(* IEC 61131-3 sources: Caravan/Archiv/12-04-19/Stations/MachineControl/MachineControl/Network/HW_Network, 1 file *)

(* ---- ONE_HW_Network_Table.st ---- *)
#define OBJECTS_CONFIG

//Define part of class SdiasBase
//Address to access the Dataobject list via SPI SDO Read
#define SDIAS_SPI_DATA_OBJECT_LIST_PAGE_ADDRESS 16#FFFF
#define SDIAS_SPI_DATA_OBJECT_LIST_PAGE_OFFSET 16#00
#define SDIAS_SPI_DATA_OBJECT_LIST_IDENTIFIER 16#12345678

//Defines the number of optional list elements in the SPI List

#define SDIAS_SPI_NUMBER_OF_OPTIONAL_ELEMENTS 7

//#pragma message("EisMic 27.06.2014 14:44 \ Noch schauen ob ichs besser machen kann")
#define SDIAS_SPI_HEADER_BEFORE_OPTIONAL_ELEMENTS 16#18
#define SDIAS_SPI_HARDWARE_VERSION_OFFSET 16#C
#define SDIAS_SPI_VENDOR_ID_OFFSET 16#0

//SPI List IDs
#define SDIAS_SPI_IDENTIFICATION_LIST_ID 1
#define SDIAS_SPI_FLASH_CONFIGURATION_ID 2
#define SDIAS_SPI_VENDOR_NAME_ID 3
#define SDIAS_SPI_DEVICE_NAME_ID 4
#define SDIAS_SPI_SERIAL_NUMBER_ID 5
#define SDIAS_SPI_ORDERING_NUMBER_ID 6
#define SDIAS_SPI_DOCUMENTATION_PDF_ID 7
#define SDIAS_SPI_CALIB_DATA_ID 10
#define SDIAS_SPI_PDO_INFORMATION_ID 128
#include "..\..\Class\SdiasManager\SdiasManager.h"
#include "..\..\Class\SdiasBase\SdiasBase.h"
#include "..\..\Class\HwControl\HwControl.h"
#include "..\..\Source\interfaces\lsl_st_hardwaretree.h"
#include "..\..\Source\interfaces\lsl_st_mt.h"
//Define part of class AI075
#define DEVICE_ID_AI075 1007

#define AI075_ADDR_CYC_WRITE        16#000
#define AI075_ADDR_CYC_READ         16#080
#define AI075_ADDR_CFG_FIRMWARE     16#100
#define AI075_ADDR_STATE_FIRMWARE   16#180

#define AI075_SDO_RESPONSE_TIMEOUT  SDIAS_SDO_TIMEOUT * 2

#define AI075_LENGTH_STATE_FIRMWARE 2
#define AI075_NUMBER_OF_ANALOG_IN   6
#define AI075_NUMBER_OF_TMP_IN      1
#define AI075_INVALID_VALUE         16#80000010$DINT
#define AI075_CABLE_BREAK_MASK      16#7F  //7 BITS
#define AI075_SHORT_CIRCUIT_MASK    16#03  //2 BITS
#define AI075_SAMPLE_POINT_MASK     16#0F  //4 BITS
#define AI075_OFFSET_SAMPLE_POINT_BITS 11

#define AI075_FIRMWARE_MIN          -10000
#define AI075_FIRMWARE_MAX          10000

//Sample Point Defines
//**************************************************************
#define AI075_FIRMWARE_VERSION_SAMPLE_POINTS_AVAILABLE  16#200
#define AI075_SAMPLE_POINTS_OFFSET_AFTER_SYNC   15    //Minimal offset that a sample point can be set after sync
#define AI075_SAMPLE_POINTS_OFFSET_BEFORE_SYNC  162   //Maximal offset that a sample point can be before next sync
//Define part of class AI088
#define DEVICE_ID_AI088 1009

#define AI088_ADDR_CYC_WRITE        16#000
#define AI088_ADDR_CYC_READ         16#080
#define AI088_ADDR_CFG_FIRMWARE     16#100
#define AI088_ADDR_STATE_FIRMWARE   16#180

#define AI088_SDO_RESPONSE_TIMEOUT  SDIAS_SDO_TIMEOUT * 2

#define AI088_LENGTH_STATE_FIRMWARE 2
#define AI088_NUMBER_OF_TMP_INPUT   10
#define AI088_CABLE_BREAK_MASK      16#3FF  //10 BITS
#define AI088_SHORT_CIRCUIT_MASK    16#3    //2 BITS
#define AI088_INVALID_VALUE         16#80000010$DINT

#define AI088_FIRMWARE_VERSION_INT_TEMP_REF 16#200  //Firmware version since when internal temperature reference and message counter are supported
#define AI088_HARDWARE_VERSION_INT_TEMP_REF 16#300  //Hardware version since when internal temperature reference are supported
// for TMP_XSelect = 10: data coming from FW may be originally negative but are
// sent as UINT type - so negativ values are sent as very big UINT values
// values greater than AI088_THRESHOLD_NEG_VALS are interpreted as neative ones
#define AI088_THRESHOLD_NEG_VALS  59000
#define AI088_SUBTRACT_FOR_INT    16#10000
//Define part of class BusInterfaceSDIASInternal
#define BUSIF_INTERNAL_MAX_NR_DO 100

// Defines for Mutex Generation
#define INTERNAL_STR_MUTEX_NAME_SEPERATOR ".."
#define INTERNAL_MUTEX_NAME_END_LENGTH 5
#define INTERNAL_MUTEX_NAME_MAX_LENGTH 32
#include "..\..\Source\BusInterface.h"
//Define part of class DI203
#define DEVICE_ID_DI203 1018
#include "..\..\Class\HwControl\watchdog.h"
#include "..\..\Source\interfaces\lsl_st_sysinfo.h"
#include "..\..\Source\interfaces\lsl_st_systrace.h"
#include <.\lsl_st_mt.h>
//Define part of class SafetyUDP
#define SAFETY_UDP_MAX_SOCKETS                6     // Max number of socket

#define SAFETY_UDP_CLT_SEND_OK                0    // Send ok
#define SAFETY_UDP_CLT_INVALID_HANDLE        -1    // Invalid handle
#define SAFETY_UDP_CLT_NOT_OPEN              -2    // Socket is not open
#define SAFETY_UDP_CLT_SEND_FAILED           -3    // Send failed
#define SAFETY_UDP_CLT_SEND_BUFFER_FULL      -4    // Send buffer is full
#define SAFETY_UDP_CLT_DATA_TO_BIG           -5    // Data to big

#define SAFETY_UDP_MAXIMUM_SEGMENT_SIZE    1452    // Maximum of user data

#define SAFETY_UDP_TIMEOUT_OPENSOCKET    (1000)    //timeout for opening socket

#define SAFETY_UDP_RECEIVE_TIMEOUT          800

#define SAFETY_UDP_TX_BUFFER_SIZE          1024
//Define part of class SafetyManager
#define LogBufferSize 1000
#include "..\..\Class\SafetyManager\SafetyManager.h"
#include "..\..\Source\interfaces\lsl_st_safetydll.h"
//Define part of class SdiasManager
#define SDIAS_SDO_MAX_LENGTH              128
#define SDIAS_SDO_RINGBUFFER_NO            64
#define SDIAS_SDO_CHANNEL_NO                3   // fixed in the VI hardware to be 3

// watchdog trigger interval (after 130ms of no trigger the SDIAS HW goes into reset again and takes at least another 10ms to be ready again)
#define SDIAS_WATCHDOG_TRIGGER_TIME        40

// time needed by sdias modules to start up after the watchdog is triggered the first time in ms
#define SDIAS_HARDWARE_STARTUP_TIME        15

// sdias manager needs 2 ticks to handle event for read task (measure sync time)
#define SDIAS_SYNC_MEASURE_TICKS            2

// after activating the PLL SyncOut it takes 3 cycles until the SDIAS sync can be injected
#define SDIAS_CYCLES_WAIT_AFTER_SYNC_ENABLE 3

// wait 1 bus cycle at start to get valid numbers in the task info
#define SDIAS_TASKINFO_READY_TICKS          1

// time to wait (in ms) until other tasks in the same or lower priority than post init have done their stuff
#define SDIAS_WAIT_TIME_IN_POST_INIT        1

#define SIZE_PER_SDIAS_CLIENT               16#0400

// for far memory accesses: 1 module can hold maximum 256 1K blocks (0-255)
#define SDIAS_1K_BLOCK_NO                       256

// far memory accesses maximum length in bytes
#define SDIAS_MAX_SIZE_FAR_MEM_ACCESS           127

#define SDIAS_OFFSET_HW_CONFIG              16#FF00
#define SDIAS_OFFSET_TASK_EVENT_IDS         16#FF10
#define SDIAS_OFFSET_FEATURE_INFO           16#FF18
#define SDIAS_OFFSET_APPLI_LED_STATES       16#FF20
#define SDIAS_OFFSET_SYNC_INJECTION_CFG     16#FF3D
#define SDIAS_OFFSET_TRIGGER_UNIT_SETUP_0   16#FF41
#define SDIAS_OFFSET_TRIGGER_UNIT_SETUP_1   16#FF45
#define SDIAS_OFFSET_TASK_START_CFG_0       16#FF60
#define SDIAS_OFFSET_TASK_CONFIG_0          16#FF86
#define SDIAS_OFFSET_TASK_CONFIG_1          16#FF96
#define SDIAS_OFFSET_TASK_INFO_1            16#FF94
#define SDIAS_OFFSET_TASK_HANDSHAKE_1       16#FF9B
#define SDIAS_OFFSET_TASK_DURATION_TIME_1   16#FF9C
#define SDIAS_OFFSET_TASK_DURATION_TIME_2   16#FFAC
#define SDIAS_OFFSET_TASK_CONFIG_2          16#FFA6

#define SDIAS_RETRIES_ALLOWED         2

// mask to get global error flag out of message counter byte of SDO responses
#define SDIAS_MASK_GLOBAL_ERROR_FLAG        16#80

// mask to get message counter out of message counter byte of SDO responses
#define SDIAS_MASK_MESSAGE_COUNTER          16#3F

#define SDIAS_EVENT_MASK_ID_SYNC_OUT0       16#10
#define SDIAS_EVENT_MASK_ID_SYNC_OUT1       16#11
#define SDIAS_EVENT_MASK_ID_SYNC_OUT2       16#12
#define SDIAS_EVENT_MASK_ID_SYNC_OUT3       16#13

#define SDIAS_MANAGER_SYNC_SYNCOUT_ID       16#85
#define SDIAS_TASK_START_EVENT_SYNCOUT_ID   16#86

#define SDIAS_PLACE_NO_MODULE_ADDED_SO_FAR  16#80000000

#define SDIAS_TRIGGER_UNIT_BYTE_SIZE        2

#define SDIAS_WAIT_TIME_FIRMWARE_HANDSHAKE  5 * 1000

// if the firmware version is below this, there might be problems with SCP111 and other modules => print warning at startup
#define SDIAS_FW_VERSION_SDO_ERROR_FIXED    16#120

// if the protocol version ist below this, Control Read/Broadcast Write Command is not supported by sdiasmanager
#define SDIAS_PROTOCOLVERSION_BROADCAST     16#120

// if the cil version ist below this, Control Read/Broadcast Write Command is not supported by OS for local SDIAS.
#define SDIAS_CILVERSION_BROADCAST         16#5001

// timeout for blocking the init during initialisation (in ms)
#define SDIAS_INIT_BLOCK_TIMEOUT            20 * 1000

#define SDIAS_MUTEX_NAME_END_LENGTH 3
#define SDIAS_MUTEX_NAME_MAX_LENGTH 32
#define SDIAS_MUTEX_STR_SEPERATOR   ".."

//#define SDIAS_RT_TIME_MEASUREMENT
#ifdef SDIAS_RT_TIME_MEASUREMENT
  #pragma message("ATTENTION: SDIAS real time measurement is active and needs additional ressources in the realtime task")
#endif

(* SDIAS data object commands  *)
#define	 SDIAS_CMD_END							  0x00			(* End command										          *)
#define	 SDIAS_CMD_ACC_MEMORY				  0x01			(* Access dpram memory								      *)
#define	 SDIAS_CMD_ACC_CONTROL				0x02			(* Access dpram control memory						  *)
#define	 SDIAS_CMD_GLOBAL						  0x03			(* SDIAS global command								      *)
#define	 SDIAS_CMD_COPY_LOCAL					0x04			(* DPRAM copy command in local dpram				*)
#define	 SDIAS_CMD_JMP_LOCAL					0x05			(* DPRAM jump command in local dpram 				*)
#define  SDIAS_CMD_ACC_MEMORY_FAR     0x07      (* SDIAS Far Memory Access                  *)

(* SDIAS defines for data object handling *)
// Write data oject list
#define	 SDIAS_DOL_WRITE_USAGE_DOL_EMPTY	  0x20			(* Usage of empty write dol list (wachtdog trigger + end command)   *)
#define	 SDIAS_DOL_WRITE_USAGE_DTA_EMPTY	  0x03			(* Usage of empty write dol data (DO ctrl of 2x copy command for task information + DO ctrl of watchdog trigger      *)
#define	 SDIAS_DOL_WRITE_OFFSET_END_CMD			0x10			(* One data object in list - offset = 1 DO size = 0x10						  *)
#define	 SDIAS_DOL_WRITE_OFFSET_FIRST_DTA		0x02			(* Offset of first data byte of second copy command = 2 (DO ctrl)   *)
#define	 SDIAS_DOL_WRITE_OFFSET_LAST_DTA		0x02			(* Offset of last data byte of second copy command = 2 (DO ctrl )   *)

// Read data oject list
#define	 SDIAS_DOL_READ_USAGE_DOL_EMPTY	    0x30			(* Usage of empty read dol list (2x task info copy command + end command)   *)
#define	 SDIAS_DOL_READ_USAGE_DTA_EMPTY	    0x0D			(* Usage of empty write dol data (DO ctrl of 2x copy command for task information + DO ctrl of watchdog trigger      *)
#define	 SDIAS_DOL_READ_OFFSET_END_CMD			0x20			(* One data object in list - offset = 1 DO size = 0x10						          *)
#define	 SDIAS_DOL_READ_OFFSET_FIRST_DTA		0x07			(* Offset of first data byte of second copy command = 7 = DO state          *)
#define	 SDIAS_DOL_READ_OFFSET_LAST_DTA		  0x0C			(* Offset of last data byte of second copy command = 12 (last byte of task information)       *)

//Versionsnumber where SDIAS SPI Read Accesses are available
#define  SDIAS_SDO_SPI_FIRMWARE_VERSION_AVAILABLE 16#0120

//error info mask
#define  SDIAS_ERROR_INFO_MASK    2#1000011000011111

// Broadcast DO Info
#define SDIAS_OFFSET_CLIENT_CTRLTIMESTAMP   16#0190
#define SDIAS_NR_TIMEBROADCAST_DOS 2
#define SDIAS_TIMEBROADCAST_SUBCMD 16#B0
#include "..\..\Source\interfaces\lsl_st_pll.h"
//Define part of class SdiasPLC
#define SDIASM_OBJECT_PATH            16#88000002   // Object Path for VSDIASmanager Length = 2 (First 2byte), Domain = 0 (3rd byte), Escape Sequence SDIAS (4th byte)
//Define part of class SR020
#define DEVICE_ID_SR020             1015        //DeviceID of SR020

#define SR020_ADDR_CYC_WRITE        16#00       //Address for TPDO
#define SR020_ADDR_CYC_READ         16#0A       //Address for RPDO

#define SR020_ADDR_CFG_FIRMWARE     16#200      //Address-Offset to the Configuration of the Firmware
#define SR020_ADDR_STATE_FIRMWARE   16#280      //Address-Offset to the Status of the Firmware
#define SR020_ADDR_I2T_THRESHOLD    16#20       //Address-Offset to Write I²T Threshold
#define SR020_ADDR_LED_MAX          16#18       //Address-Offset to get LED Configuration-Values

//Define for the H-Brdige
//-----------------------------------------------------------
#define SR020_GATE_A_LOW		          2#0100000000000000    //Bit-Configuration for Enable GateA Low-Switch
#define SR020_GATE_A_HIGH		          2#0001000000000000    //Bit-Configuration for Enable GateA High-Switch
#define SR020_GATE_B_LOW		          2#1000000000000000    //Bit-Configuration for Enable GateB Low-Switch
#define SR020_GATE_B_HIGH		          2#0010000000000000    //Bit-Configuration for Enable GateB High-Switch

#define SR020_MASK_CONTROL	          16#0FFF     //Mask for Output Sequence Bits
#define SR020_MASK_TIME		            16#F000     //Mask for TimeValue

#define SR020_T_SWITCH                41      //Delay Time for Switch
#define SR020_DEFAULT_SEQ_INIT        1       //Initilization for Sequencer => After 1 FPGA-Cycle switch to next Sequency

#define SR020_FPGA_FREQ_MHZ           50    //Frequency of FPGA

#define SR020_SDO_RESPONSE_TIMEOUT  SDIAS_SDO_TIMEOUT * 2     //SDO-Response Timeout

//#define SR020_I2T_THRESHOLD          16000000   //Maximal allowed I²T Value in mA²s ==> 16 A²s
//#pragma message ("TarPet: dieser Wert wurde vorest empirisch ermittelt und sollte noch genau bestimmt werden");
#define SR020_I2T_THRESHOLD          78000   //Maximal allowed I²T Value in mA²s ==> 16 A²s

#define SR020_SPEED_SCALING          10000      //Scaling of the Server Speed (0.00% to 100.00%)
#define SR020_MINPULSE_SCALING       1000       //Scaling of the Server MinPulse (0.0% to 100.0%)

#define SR020_STATUS_BITS_LATCHED  2#0001110011110 // no DC OK info, no sequencer info, no Overtemperature and no I2C error
#define SR020_STATUS_BITS          2#1010000000000 // Overtemperature and I2C error
#define SR020_STATUS_BITS_INVERTED 2#0000001100001 // DC OK info and sequencer info
//Define part of class TO161
#define DEVICE_ID_TO161 1004

#define TO161_ADDR_CYC_WRITE  0
#define TO161_ADDR_CYC_READ   2

#define TO161_WRITE_LENGTH    2
#define TO161_READ_LENGTH     2

FUNCTION GLOBAL TAB ONE_HW_Network
-1$UINT, 0$UINT,
0$UINT, 0$UINT,

24$UDINT,
TO_UDINT(529317953), "_CanLib", 1$UINT, 10$UINT, 2$UINT,
TO_UDINT(4078275645), "_SerLib", 1$UINT, 34$UINT, 2$UINT,
TO_UDINT(2809270484), "AI075", 1$UINT, 36$UINT, 1$UINT,
TO_UDINT(1583050918), "AI088", 1$UINT, 34$UINT, 1$UINT,
TO_UDINT(3882880897), "BusInterfaceSDIASInternal", 2$UINT, 0$UINT, 0$UINT,
TO_UDINT(3961086008), "CP102_IOs", 1$UINT, 0$UINT, 1$UINT,
TO_UDINT(794617671), "CriticalSection", 0$UINT, 4$UINT, 2$UINT,
TO_UDINT(3392436280), "DI203", 1$UINT, 30$UINT, 1$UINT,
TO_UDINT(2471641665), "HwControl", 5$UINT, 2$UINT, 1$UINT,
TO_UDINT(1193052171), "HwControlBase", 1$UINT, 10$UINT, 0$UINT,
TO_UDINT(4260294091), "HWRtPostScan", 1$UINT, 0$UINT, 1$UINT,
TO_UDINT(2225119864), "MerkerEx", 1$UINT, 22$UINT, 5$UINT,
TO_UDINT(1799751072), "SafetyManager", 2$UINT, 11$UINT, 1$UINT,
TO_UDINT(3727715967), "SafetyUDP", 1$UINT, 2$UINT, 0$UINT,
TO_UDINT(3175101883), "SdiasBase", 1$UINT, 58$UINT, 0$UINT,
TO_UDINT(4173303375), "SdiasHubBase", 1$UINT, 10$UINT, 1$UINT,
TO_UDINT(2118381352), "SdiasManager", 1$UINT, 92$UINT, 1$UINT,
TO_UDINT(1159122596), "SdiasPLC", 2$UINT, 0$UINT, 1$UINT,
TO_UDINT(928449634), "SR020", 1$UINT, 34$UINT, 1$UINT,
TO_UDINT(1850111279), "String", 1$UINT, 10$UINT, 5$UINT,
TO_UDINT(2898603620), "StringInternal", 1$UINT, 82$UINT, 0$UINT,
TO_UDINT(900581525), "TO161", 1$UINT, 32$UINT, 1$UINT,
TO_UDINT(3232495061), "VirtualBaseInit", 1$UINT, 3$UINT, 0$UINT,
TO_UDINT(819479645), "XXXBase_IOs", 1$UINT, 0$UINT, 0$UINT,

1$UINT, TO_UDINT(2156319869), "CP102_IOS2\_BASE\_CANLIB1",
1$UINT, TO_UDINT(428836295), "CP102_IOS2\_BASE\_CANLIB2",

1$UINT, TO_UDINT(3654905894), "CP102_IOS2\_BASE\_SERLIB1",
1$UINT, TO_UDINT(1087381916), "CP102_IOS2\_BASE\_SERLIB2",

_NO_ATTR, TO_UDINT(46500714), "AI0751",

_NO_ATTR, TO_UDINT(3157766682), "AI0881",

_NO_ATTR, TO_UDINT(842735603), "CP102_IOS2",

1$UINT, TO_UDINT(2972590922), "HWCONTROL1\SAFETYMANAGER\UDPRECEIVEDATA",
1$UINT, TO_UDINT(1868223583), "HWCONTROL1\SAFETYMANAGER\UDPSENDDATA",

_NO_ATTR, TO_UDINT(2870240081), "DI2031",

_NO_ATTR, TO_UDINT(2190789875), "HWCONTROL1",

1$UINT, TO_UDINT(1673205898), "HWCONTROL1\HWRTPOSTSCAN",

1$UINT, TO_UDINT(588388748), "AI0751\_BASE\SERIALNOSTR\MERKEREX0",
1$UINT, TO_UDINT(2299507738), "AI0881\_BASE\SERIALNOSTR\MERKEREX0",
1$UINT, TO_UDINT(212455792), "DI2031\_BASE\SERIALNOSTR\MERKEREX0",
1$UINT, TO_UDINT(1493349760), "SR0201\_BASE\SERIALNOSTR\MERKEREX0",
1$UINT, TO_UDINT(146675376), "TO1611\_BASE\SERIALNOSTR\MERKEREX0",

1$UINT, TO_UDINT(1778590035), "HWCONTROL1\SAFETYMANAGER",

1$UINT, TO_UDINT(1007630054), "SDIASPLC1\SDIASHUBBASE1",

1$UINT, TO_UDINT(4015996540), "SDIASPLC1\SDIASMANAGER1",

_NO_ATTR, TO_UDINT(1378000520), "SDIASPLC1",

_NO_ATTR, TO_UDINT(542619847), "SR0201",

1$UINT, TO_UDINT(1502199223), "AI0751\_BASE\SERIALNOSTR",
1$UINT, TO_UDINT(2748134452), "AI0881\_BASE\SERIALNOSTR",
1$UINT, TO_UDINT(1916703938), "DI2031\_BASE\SERIALNOSTR",
1$UINT, TO_UDINT(777954792), "SR0201\_BASE\SERIALNOSTR",
1$UINT, TO_UDINT(3843311503), "TO1611\_BASE\SERIALNOSTR",

_NO_ATTR, TO_UDINT(59516340), "TO1611",

//Internal connections
0$UDINT,
20$UDINT,
TO_UDINT(4), "SerialNoStr", TO_UDINT(22),
TO_UDINT(5), "SerialNoStr", TO_UDINT(23),
TO_UDINT(6), "_SerLib1", TO_UDINT(2),
TO_UDINT(6), "_SerLib2", TO_UDINT(3),
TO_UDINT(6), "_CanLib1", TO_UDINT(0),
TO_UDINT(6), "_CanLib2", TO_UDINT(1),
TO_UDINT(9), "SerialNoStr", TO_UDINT(24),
TO_UDINT(10), "SafetyManager", TO_UDINT(17),
TO_UDINT(10), "HWRtPostScan", TO_UDINT(11),
TO_UDINT(17), "UdpSendData", TO_UDINT(8),
TO_UDINT(17), "UdpReceiveData", TO_UDINT(7),
TO_UDINT(20), "SdiasManager1", TO_UDINT(19),
TO_UDINT(20), "SdiasHubBase1", TO_UDINT(18),
TO_UDINT(21), "SerialNoStr", TO_UDINT(25),
TO_UDINT(22), "MerkerEx0", TO_UDINT(12),
TO_UDINT(23), "MerkerEx0", TO_UDINT(13),
TO_UDINT(24), "MerkerEx0", TO_UDINT(14),
TO_UDINT(25), "MerkerEx0", TO_UDINT(15),
TO_UDINT(26), "MerkerEx0", TO_UDINT(16),
TO_UDINT(27), "SerialNoStr", TO_UDINT(26),
0$UDINT,
16$UDINT,
TO_UDINT(4), "SdiasIn", TO_UDINT(18), "ClassSvr",
TO_UDINT(5), "SdiasIn", TO_UDINT(18), "ClassSvr",
TO_UDINT(6), "To_HwControl", TO_UDINT(10), "Control",
TO_UDINT(9), "SdiasIn", TO_UDINT(18), "ClassSvr",
TO_UDINT(11), "toHwControlBase", TO_UDINT(10), "Control",
TO_UDINT(17), "To_HwControl", TO_UDINT(10), "Control",
TO_UDINT(18), "ToNextSDIAS", TO_UDINT(19), "ClassState",
TO_UDINT(19), "ToBusInterface", TO_UDINT(20), "CallCommand",
TO_UDINT(20), "ToHwControl", TO_UDINT(10), "Control",
TO_UDINT(21), "SdiasIn", TO_UDINT(18), "ClassSvr",
TO_UDINT(22), "DataBuffer", TO_UDINT(12), "m_udLength",
TO_UDINT(23), "DataBuffer", TO_UDINT(13), "m_udLength",
TO_UDINT(24), "DataBuffer", TO_UDINT(14), "m_udLength",
TO_UDINT(25), "DataBuffer", TO_UDINT(15), "m_udLength",
TO_UDINT(26), "DataBuffer", TO_UDINT(16), "m_udLength",
TO_UDINT(27), "SdiasIn", TO_UDINT(18), "ClassSvr",

//Initialization values
0$UDINT,
67$UDINT,
TO_UDINT(0), "CanBus", TO_UDINT(0),//|HW_Network._base\CP102_IOs2\_CanLib1.CanBus;
TO_UDINT(1), "CanBus", TO_UDINT(1),//|HW_Network._base\CP102_IOs2\_CanLib2.CanBus;
TO_UDINT(2), "Com", TO_UDINT(0),//|HW_Network._base\CP102_IOs2\_SerLib1.Com;
TO_UDINT(3), "Com", TO_UDINT(1),//|HW_Network._base\CP102_IOs2\_SerLib2.Com;
TO_UDINT(4), "LEDControl", TO_UDINT(0),//|HW_Network.AI0751.LEDControl;
TO_UDINT(4), "ActivateSamplePointConfig", TO_UDINT(0),//|HW_Network.AI0751.ActivateSamplePointConfig;
TO_UDINT(4), "Place", TO_UDINT(0),//|HW_Network.AI0751.Place;
TO_UDINT(4), "Required", TO_UDINT(1),//|HW_Network.AI0751.Required;
TO_UDINT(4), "AI1_Min", TO_UDINT(-10000),//|HW_Network.AI0751.AI1_Min;
TO_UDINT(4), "AI1_Max", TO_UDINT(10000),//|HW_Network.AI0751.AI1_Max;
TO_UDINT(4), "AI2_Min", TO_UDINT(-10000),//|HW_Network.AI0751.AI2_Min;
TO_UDINT(4), "AI2_Max", TO_UDINT(10000),//|HW_Network.AI0751.AI2_Max;
TO_UDINT(4), "AI3_Min", TO_UDINT(-10000),//|HW_Network.AI0751.AI3_Min;
TO_UDINT(4), "AI3_Max", TO_UDINT(10000),//|HW_Network.AI0751.AI3_Max;
TO_UDINT(4), "AI4_Min", TO_UDINT(-10000),//|HW_Network.AI0751.AI4_Min;
TO_UDINT(4), "AI4_Max", TO_UDINT(10000),//|HW_Network.AI0751.AI4_Max;
TO_UDINT(4), "AI5_Min", TO_UDINT(-10000),//|HW_Network.AI0751.AI5_Min;
TO_UDINT(4), "AI5_Max", TO_UDINT(10000),//|HW_Network.AI0751.AI5_Max;
TO_UDINT(4), "AI6_Min", TO_UDINT(-10000),//|HW_Network.AI0751.AI6_Min;
TO_UDINT(4), "AI6_Max", TO_UDINT(10000),//|HW_Network.AI0751.AI6_Max;
TO_UDINT(4), "UseSamplePointConfig", TO_UDINT(0),//|HW_Network.AI0751.UseSamplePointConfig;
TO_UDINT(5), "LEDControl", TO_UDINT(0),//|HW_Network.AI0881.LEDControl;
TO_UDINT(5), "Place", TO_UDINT(4),//|HW_Network.AI0881.Place;
TO_UDINT(5), "Required", TO_UDINT(1),//|HW_Network.AI0881.Required;
TO_UDINT(5), "TMP_1Select", TO_UDINT(10),//|HW_Network.AI0881.TMP_1Select;
TO_UDINT(5), "TMP_1RefSensor", TO_UDINT(0),//|HW_Network.AI0881.TMP_1RefSensor;
TO_UDINT(5), "TMP_2Select", TO_UDINT(10),//|HW_Network.AI0881.TMP_2Select;
TO_UDINT(5), "TMP_2RefSensor", TO_UDINT(0),//|HW_Network.AI0881.TMP_2RefSensor;
TO_UDINT(5), "TMP_3Select", TO_UDINT(1),//|HW_Network.AI0881.TMP_3Select;
TO_UDINT(5), "TMP_3RefSensor", TO_UDINT(0),//|HW_Network.AI0881.TMP_3RefSensor;
TO_UDINT(5), "TMP_4Select", TO_UDINT(1),//|HW_Network.AI0881.TMP_4Select;
TO_UDINT(5), "TMP_4RefSensor", TO_UDINT(0),//|HW_Network.AI0881.TMP_4RefSensor;
TO_UDINT(5), "TMP_5Select", TO_UDINT(1),//|HW_Network.AI0881.TMP_5Select;
TO_UDINT(5), "TMP_5RefSensor", TO_UDINT(0),//|HW_Network.AI0881.TMP_5RefSensor;
TO_UDINT(5), "TMP_6RefSensor", TO_UDINT(0),//|HW_Network.AI0881.TMP_6RefSensor;
TO_UDINT(5), "TMP_7RefSensor", TO_UDINT(0),//|HW_Network.AI0881.TMP_7RefSensor;
TO_UDINT(5), "TMP_8RefSensor", TO_UDINT(0),//|HW_Network.AI0881.TMP_8RefSensor;
TO_UDINT(9), "LEDControl", TO_UDINT(0),//|HW_Network.DI2031.LEDControl;
TO_UDINT(9), "Place", TO_UDINT(1),//|HW_Network.DI2031.Place;
TO_UDINT(9), "Required", TO_UDINT(1),//|HW_Network.DI2031.Required;
TO_UDINT(10), "UdpSafetyPort", TO_UDINT(10823),//|HW_Network.HwControl1.UdpSafetyPort;
TO_UDINT(10), "InterfaceNo", TO_UDINT(1),//|HW_Network.HwControl1.InterfaceNo;
TO_UDINT(12), "ThreadSafe", TO_UDINT(0),//|HW_Network.SerialNoStr\_base\AI0751\MerkerEx0.ThreadSafe;
TO_UDINT(13), "ThreadSafe", TO_UDINT(0),//|HW_Network.SerialNoStr\_base\AI0881\MerkerEx0.ThreadSafe;
TO_UDINT(14), "ThreadSafe", TO_UDINT(0),//|HW_Network.SerialNoStr\_base\DI2031\MerkerEx0.ThreadSafe;
TO_UDINT(15), "ThreadSafe", TO_UDINT(0),//|HW_Network.SerialNoStr\_base\SR0201\MerkerEx0.ThreadSafe;
TO_UDINT(16), "ThreadSafe", TO_UDINT(0),//|HW_Network.SerialNoStr\_base\TO1611\MerkerEx0.ThreadSafe;
TO_UDINT(17), "UdpSafetyPort", TO_UDINT(10823),//|HW_Network.HwControl1\SafetyManager.UdpSafetyPort;
TO_UDINT(17), "InterfaceNo", TO_UDINT(1),//|HW_Network.HwControl1\SafetyManager.InterfaceNo;
TO_UDINT(18), "SplitterPlace", TO_UDINT(0),//|HW_Network.SdiasPLC1\SdiasHubBase1.SplitterPlace;
TO_UDINT(19), "DeviceID", TO_UDINT(0),//|HW_Network.SdiasPLC1\SdiasManager1.DeviceID;
TO_UDINT(20), "CycleTime", TO_UDINT(1000),//|HW_Network.SdiasPLC1.CycleTime;
TO_UDINT(20), "IsoStartPoint", TO_UDINT(50),//|HW_Network.SdiasPLC1.IsoStartPoint;
TO_UDINT(21), "LEDControl", TO_UDINT(0),//|HW_Network.SR0201.LEDControl;
TO_UDINT(21), "MinPulse", TO_UDINT(7),//|HW_Network.SR0201.MinPulse;
TO_UDINT(21), "Place", TO_UDINT(3),//|HW_Network.SR0201.Place;
TO_UDINT(21), "Required", TO_UDINT(1),//|HW_Network.SR0201.Required;
TO_UDINT(21), "PWMPeriod", TO_UDINT(32),//|HW_Network.SR0201.PWMPeriod;
TO_UDINT(21), "I2TThreshold", TO_UDINT(100),//|HW_Network.SR0201.I2TThreshold;
TO_UDINT(22), "SingleRealloc", TO_UDINT(1),//|HW_Network._base\AI0751\SerialNoStr.SingleRealloc;
TO_UDINT(23), "SingleRealloc", TO_UDINT(1),//|HW_Network._base\AI0881\SerialNoStr.SingleRealloc;
TO_UDINT(24), "SingleRealloc", TO_UDINT(1),//|HW_Network._base\DI2031\SerialNoStr.SingleRealloc;
TO_UDINT(25), "SingleRealloc", TO_UDINT(1),//|HW_Network._base\SR0201\SerialNoStr.SingleRealloc;
TO_UDINT(26), "SingleRealloc", TO_UDINT(1),//|HW_Network._base\TO1611\SerialNoStr.SingleRealloc;
TO_UDINT(27), "LEDControl", TO_UDINT(0),//|HW_Network.TO1611.LEDControl;
TO_UDINT(27), "Place", TO_UDINT(2),//|HW_Network.TO1611.Place;
TO_UDINT(27), "Required", TO_UDINT(1),//|HW_Network.TO1611.Required;

//Symbolic initialization values
0$UDINT,
0$UDINT,

//Initialization of string values
0$UDINT,
0$UDINT,

//Configuration of tasks (RealTime, Cyclic, Background)
0$UDINT,
1$UDINT,
TO_UDINT(11), (1)$UDINT, 4194304$DINT, 	//HWCONTROL1\HWRTPOSTSCAN

0$UDINT,
0$UDINT,

0$UDINT,
0$UDINT,

//External connections
0$UDINT,
0$UDINT,

//Magic internal connections
0$UDINT,
3$UDINT,
TO_UDINT(17), "UdpSafetyPort", TO_UDINT(10), "UdpSafetyPort",
TO_UDINT(17), "InterfaceNo", TO_UDINT(10), "InterfaceNo",
TO_UDINT(17), "SafetyDomainTimeout", TO_UDINT(10), "SafetyDomainTimeout",

//Configuration of timeslots of tasks (RealTime, Cyclic)
#ifdef __LSLLDR_TIMESLOTS__
0$UDINT,
0$UDINT,

0$UDINT,
0$UDINT,

#endif //__LSLLDR_TIMESLOTS__

//MultiMaster connections
#ifdef __LSLLDR_MULTIMASTER__
0$UDINT,
0$UDINT,
#endif //__LSLLDR_MULTIMASTER__

//Configuration for task ID (RealTime, CyclicTime)
#ifdef __LSLLDR_TASKID__
"\\\\TASKS2  "
0$UDINT,
1$UDINT,
(0)$UDINT, 	//HWCONTROL1\HWRTPOSTSCAN

0$UDINT,
0$UDINT,

0$UDINT,
0$UDINT,

#endif //__LSLLDR_TASKID__

END_FUNCTION
